(*
.. note:: This is a note admonition.
   This is the second line of the first paragraph.

   - The note contains all indented body elements
     following.
   - It includes this bullet list.
*)

FUNCTION_BLOCK FB_Libdoc_SpecificNotes
VAR_INPUT
    nVarA : INT;
    nVarB : INT;
END_VAR
VAR_OUTPUT
    nSum : INT;
END_VAR
VAR
END_VAR

END_FUNCTION_BLOCK

(* stored: Version 1.1.0.1, ProductVersion 3.1.4022.18
   POU FB_Libdoc_SpecificNotes: Id {32019413-ce36-4918-8156-39d55e3cdaee}, SpecialFunc None *)
